// TIA Portal project "Closed" (V21)

(* hardware
DEVICE "PLC_Closed"  S7-1500 station
   slot 0: "Rail_0"  Rack  6ES7 590-1***0-0AA0
   slot 1: "PLC_Closed"  CPU 1516-3 PN/DP  6ES7 516-3AN02-0AB0  V2.9
      slot 3: "CPU display_1"  6ES7591-1BA00-0AA0
      slot 32768: "PROFINET interface_1"  X1
         slot 32769: "Port_1"  X1 P1
         slot 32770: "Port_2"  X1 P2
      slot 33024: "PROFINET interface_2"  X2
         slot 33025: "Port_1"  X2 P1
      slot 33280: "DP interface_1"  X3
      slot 34817: "Virtual CP interface port_1"  Virtual CP interface port  Virtual CP interface port
*)

// ===== PLC "PLC_Closed"  CPU 1516-3 PN/DP =====
// protected blocks, not shown: "Secret"

DATA_BLOCK "CallerData"   // DB1
{ S7_Optimized_Access := 'TRUE' }
VERSION : 0.1
// stored: InstanceOfName Caller
"Caller"
BEGIN
END_DATA_BLOCK

FUNCTION_BLOCK "Caller"   // FB2, SCL
TITLE = An open block that calls the protected one
{ S7_Optimized_Access := 'TRUE' }
VERSION : 0.1
   VAR_INPUT
      seed : DInt;   // Passed on
   END_VAR
   VAR_OUTPUT
      answer : DInt;   // Passed back
   END_VAR
   VAR
      inner : "Secret";   // The protected block, as a multi-instance
   END_VAR
BEGIN

    #inner(seed := #seed);
    #answer := #inner.answer;
END_FUNCTION_BLOCK